{attribute 'qualified_only'}
VAR_GLOBAL
	VTEM_IN AT %I* : ARRAY [0..2] OF WORD;
	VTEM_OUT AT %Q* : ARRAY [0..2] OF WORD;
END_VAR

(* stored: Version 1.1.0.1, ProductVersion 3.1.4024.16
   GVL GVL: Id {fca253f4-aab3-4ff2-a27d-5a09328aa443} *)
